SUBAPPLICATION Uebung_250_AX (* Grenzfrequenz des Analogeingangs messen: dasselbe Rechtecksignal an AI (I1) und PI (I2), Vergleich der Frequenzen je 1 s Torzeit *)
  (* Standard: 61499-2; Description: Copyright (c) 2026 Meisterschulen am Ostbahnhof This program and the accompanying materials are made available under the terms of the Eclipse Public License 2.0 which is available at https://www.eclipse.org/legal/epl-2.0/ SPDX-License-Identifier: EPL-2.0 *)
  (* Version 1.0, 2026-10-29, Franz Höpfinger, Meisterschulen am Ostbahnhof, initial implementation *)
  PACKAGE Uebungen;
  IMPORT logiBUS::io::AI::logiBUS_AI::AnalogInput_I1;
  IMPORT logiBUS::io::PI::logiBUS_PI::PulseInput_I2;
  (* Documentation:
  Grenzfrequenz des Analogeingangs
   Testaufbau: ein Rechtecksignal 0-10 V gleichzeitig an I1 (als AI) und I2 (als PI). Der PI zaehlt in Hardware und liefert die echte Frequenz. Der AI liefert nur alle ca. 3,2 ms einen Mittelwert (ESP32-P4, 20 kHz Continuous-Mode, 64 Samples je Block).
    - SCHMITT macht aus dem AI-Wert ein Bit (ein ab 75 %, aus unter 25 %), AI_EDGES zaehlt dessen steigende Flanken.
   - GATE (1 s) liest beide Zaehler, F_AI und F_PI sind damit direkt in Hz. SAMPLES_S zeigt, wie viele AI-Werte pro Sekunde ankommen.
   - OK ist TRUE, solange |f_AI - f_PI| <= 2 Hz. F_GRENZ merkt sich die hoechste PI-Frequenz, bei der das noch galt.
    Oberhalb der Grenze mittelt der Treiber das Rechteck zu einem Wert um 50 %, der Schmitt-Trigger schaltet nicht mehr und f_AI faellt ab. Neu messen: Programm neu starten.
  *)
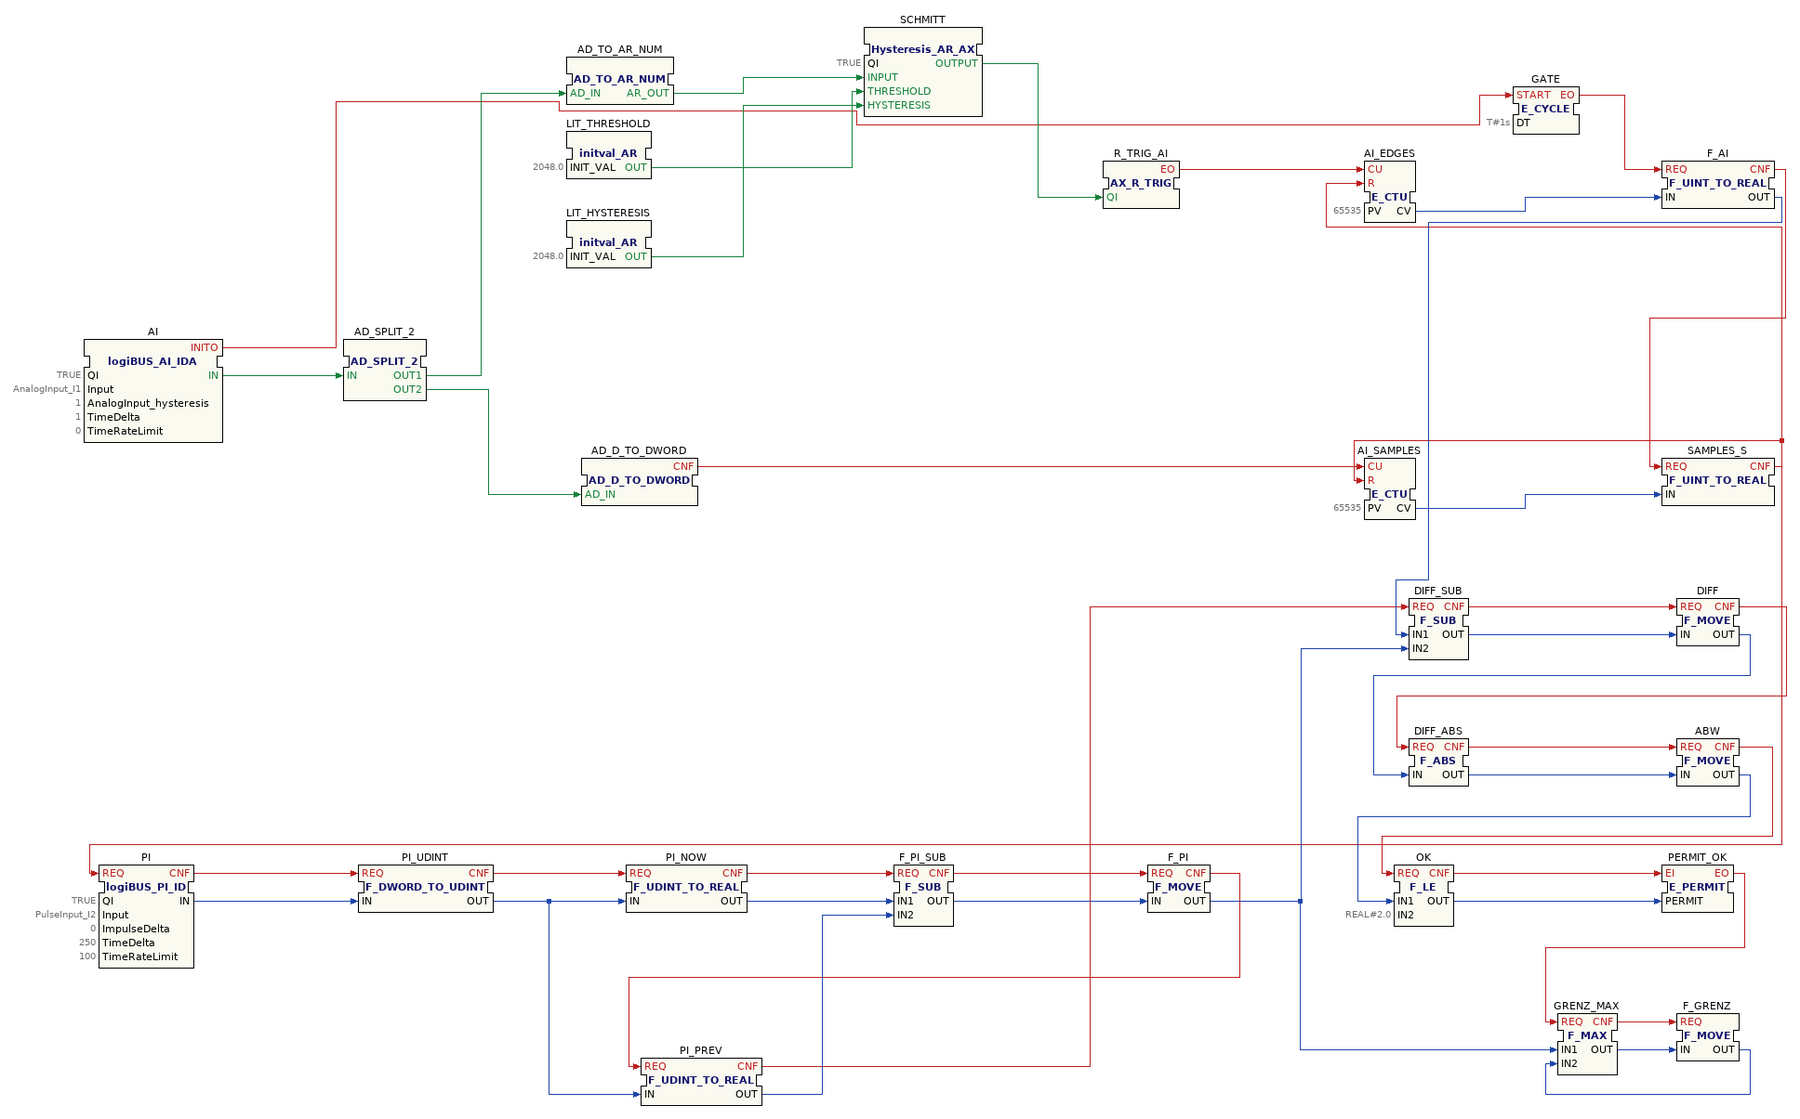
  (* Watch: F_AI.OUT, F_PI.OUT, SAMPLES_S.OUT, ABW.OUT, OK.OUT, F_GRENZ.OUT Frequenz am Generator langsam steigern. F_GRENZ.OUT = Grenzfrequenz. *)
  FBS
    AI : logiBUS::io::AI::logiBUS_AI_IDA(QI := TRUE, Input := AnalogInput_I1, AnalogInput_hysteresis := 1, TimeDelta := 1, TimeRateLimit := 0); (* Analogeingang I1, 0-10 V, jede ADC-Mittelung melden *)
    AD_SPLIT_2 : adapter::events::unidirectional::AD_SPLIT_2;
    AD_TO_AR_NUM : adapter::conversion::unidirectional::AD_TO_AR_NUM;
    LIT_THRESHOLD : adapter::types::unidirectional::AR::initval::initval_AR(INIT_VAL := 2048.0);
    LIT_HYSTERESIS : adapter::types::unidirectional::AR::initval::initval_AR(INIT_VAL := 2048.0);
    SCHMITT : logiBUS::signalprocessing::hysteresis::Hysteresis_AR_AX(QI := TRUE); (* Ein ab 3072 (75 %), aus unter 1024 (25 %) *)
    R_TRIG_AI : adapter::events::unidirectional::AX_R_TRIG;
    AI_EDGES : iec61499::events::E_CTU(PV := 65535); (* Steigende Flanken am AI je Torzeit *)
    AD_D_TO_DWORD : adapter::conversion::unidirectional::AD_D_TO_DWORD;
    AI_SAMPLES : iec61499::events::E_CTU(PV := 65535); (* AI-Werte je Torzeit (effektive Abtastrate) *)
    GATE : iec61499::events::E_CYCLE(DT := T#1s); (* Torzeit 1 s: Zaehlerstand = Frequenz in Hz *)
    F_AI : iec61131::conversion::F_UINT_TO_REAL; (* Frequenz aus AI [Hz] *)
    SAMPLES_S : iec61131::conversion::F_UINT_TO_REAL; (* AI-Werte pro Sekunde *)
    PI : logiBUS::io::PI::logiBUS_PI_ID(QI := TRUE, Input := PulseInput_I2, ImpulseDelta := 0, TimeDelta := 250, TimeRateLimit := 100); (* Pulseingang I2 als Referenz (Hardware-Zaehler) *)
    PI_UDINT : iec61131::conversion::F_DWORD_TO_UDINT;
    PI_NOW : iec61131::conversion::F_UDINT_TO_REAL;
    F_PI_SUB : iec61131::arithmetic::F_SUB;
    F_PI : iec61131::selection::F_MOVE; (* Frequenz aus PI [Hz] *) {SET_ATTRIBUTE(DataType, REAL)}
    PI_PREV : iec61131::conversion::F_UDINT_TO_REAL; (* Zaehlerstand der vorigen Torzeit *)
    DIFF_SUB : iec61131::arithmetic::F_SUB;
    DIFF : iec61131::selection::F_MOVE; (* f_AI - f_PI [Hz] *) {SET_ATTRIBUTE(DataType, REAL)}
    DIFF_ABS : iec61131::numerical::F_ABS;
    ABW : iec61131::selection::F_MOVE; (* Abweichung |f_AI - f_PI| [Hz] *) {SET_ATTRIBUTE(DataType, REAL)}
    OK : iec61131::comparison::F_LE(IN2 := REAL#2.0); (* TRUE: AI folgt dem Signal noch (Abweichung <= 2 Hz) *)
    PERMIT_OK : iec61499::events::E_PERMIT;
    GRENZ_MAX : iec61131::selection::F_MAX;
    F_GRENZ : iec61131::selection::F_MOVE; (* Grenzfrequenz: hoechste f_PI, bei der OK=TRUE war [Hz] *) {SET_ATTRIBUTE(DataType, REAL)}
  END_FBS
  EVENT_CONNECTIONS
    AI.INITO TO GATE.START;
    R_TRIG_AI.EO TO AI_EDGES.CU;
    AD_D_TO_DWORD.CNF TO AI_SAMPLES.CU;
    GATE.EO TO F_AI.REQ;
    F_AI.CNF TO SAMPLES_S.REQ;
    SAMPLES_S.CNF TO AI_EDGES.R;
    SAMPLES_S.CNF TO AI_SAMPLES.R;
    PI.CNF TO PI_UDINT.REQ;
    PI_UDINT.CNF TO PI_NOW.REQ;
    PI_NOW.CNF TO F_PI_SUB.REQ;
    F_PI_SUB.CNF TO F_PI.REQ;
    F_PI.CNF TO PI_PREV.REQ;
    PI_PREV.CNF TO DIFF_SUB.REQ;
    DIFF_SUB.CNF TO DIFF.REQ;
    DIFF.CNF TO DIFF_ABS.REQ;
    DIFF_ABS.CNF TO ABW.REQ;
    ABW.CNF TO OK.REQ;
    OK.CNF TO PERMIT_OK.EI;
    PERMIT_OK.EO TO GRENZ_MAX.REQ;
    GRENZ_MAX.CNF TO F_GRENZ.REQ;
    SAMPLES_S.CNF TO PI.REQ;
  END_CONNECTIONS
  DATA_CONNECTIONS
    AI_EDGES.CV TO F_AI.IN;
    AI_SAMPLES.CV TO SAMPLES_S.IN;
    PI.IN TO PI_UDINT.IN;
    PI_UDINT.OUT TO PI_NOW.IN;
    PI_UDINT.OUT TO PI_PREV.IN;
    PI_NOW.OUT TO F_PI_SUB.IN1;
    PI_PREV.OUT TO F_PI_SUB.IN2;
    F_PI_SUB.OUT TO F_PI.IN;
    F_AI.OUT TO DIFF_SUB.IN1;
    F_PI.OUT TO DIFF_SUB.IN2;
    DIFF_SUB.OUT TO DIFF.IN;
    DIFF.OUT TO DIFF_ABS.IN;
    DIFF_ABS.OUT TO ABW.IN;
    ABW.OUT TO OK.IN1;
    OK.OUT TO PERMIT_OK.PERMIT;
    F_PI.OUT TO GRENZ_MAX.IN1;
    F_GRENZ.OUT TO GRENZ_MAX.IN2;
    GRENZ_MAX.OUT TO F_GRENZ.IN;
  END_CONNECTIONS
  ADAPTER_CONNECTIONS
    AI.IN TO AD_SPLIT_2.IN;
    AD_SPLIT_2.OUT1 TO AD_TO_AR_NUM.AD_IN;
    AD_SPLIT_2.OUT2 TO AD_D_TO_DWORD.AD_IN;
    AD_TO_AR_NUM.AR_OUT TO SCHMITT.INPUT;
    LIT_THRESHOLD.OUT TO SCHMITT.THRESHOLD;
    LIT_HYSTERESIS.OUT TO SCHMITT.HYSTERESIS;
    SCHMITT.OUTPUT TO R_TRIG_AI.QI;
  END_CONNECTIONS
END_SUBAPPLICATION
